(* IEC 61131-3 sources: SemantiST/compiler/toolchain/compatibility/profiles/s7-conversions, 1 file *)

(* ---- conversions.st ---- *)
(* Generated by compiler/toolchain/compatibility/profiles/generate_codesys.py
   from the pinned RuSTy standard library. Do not edit by hand.
   S7-SCL conversions (S7-SCL V5.3 manual, chapter 14) on RuSTy's
   representation: DATE = days since 1990-01-01, TIME/TOD = milliseconds,
   least significant bit for INT/DINT_TO_BOOL. *)

FUNCTION INT_TO_BOOL : BOOL
VAR_INPUT IN : INT; END_VAR
VAR w : WORD; END_VAR
    w := IN;
    INT_TO_BOOL := (w AND 1) <> 0;
END_FUNCTION

FUNCTION __S7_DINT_TO_BOOL : BOOL
VAR_INPUT IN : DINT; END_VAR
VAR w : DWORD; END_VAR
    w := IN;
    __S7_DINT_TO_BOOL := (w AND 1) <> 0;
END_FUNCTION

FUNCTION DINT_TO_DATE : DATE
VAR_INPUT IN : DINT; END_VAR
VAR v : LINT; END_VAR
    v := IN;
    DINT_TO_DATE := LINT_TO_DATE((v + LINT#7305) * LINT#86400000000000);
END_FUNCTION

FUNCTION DATE_TO_DINT : DINT
VAR_INPUT IN : DATE; END_VAR
    DATE_TO_DINT := LINT_TO_DINT(DATE_TO_LINT(IN) / LINT#86400000000000 - LINT#7305);
END_FUNCTION

FUNCTION DINT_TO_TIME : TIME
VAR_INPUT IN : DINT; END_VAR
VAR v : LINT; END_VAR
    v := IN;
    DINT_TO_TIME := LINT_TO_TIME(v * LINT#1000000);
END_FUNCTION

FUNCTION TIME_TO_DINT : DINT
VAR_INPUT IN : TIME; END_VAR
    TIME_TO_DINT := LINT_TO_DINT(TIME_TO_LINT(IN) / LINT#1000000);
END_FUNCTION

FUNCTION DINT_TO_TOD : TIME_OF_DAY
VAR_INPUT IN : DINT; END_VAR
VAR v : LINT; END_VAR
    v := IN;
    DINT_TO_TOD := LINT_TO_TOD(v * LINT#1000000);
END_FUNCTION

FUNCTION TOD_TO_DINT : DINT
VAR_INPUT IN : TIME_OF_DAY; END_VAR
    TOD_TO_DINT := LINT_TO_DINT(TOD_TO_LINT(IN) / LINT#1000000);
END_FUNCTION
